// TIA Portal V19 export
// export: Created 2026-10-15T10:10:35.0564557Z, ExportSetting WithDefaults, DisplayName Totally Integrated Automation Portal, DisplayVersion V19, DisplayName TIA Portal Openness, DisplayVersion V19, DisplayName TIA Portal Version Control Interface, DisplayVersion V19, DisplayName STEP 7 Professional, DisplayVersion V19, DisplayName STEP 7 Safety, DisplayVersion V19, DisplayName WinCC Basic/Comfort/Advanced, DisplayVersion V19, DisplayName WinCC Unified, DisplayVersion V19
FUNCTION "ROLL_ShowRecipe" : Void   // FC11, SCL
{ S7_Optimized_Access := 'TRUE' }
VERSION : 0.1
// stored: AutoNumber true, IsIECCheckEnabled false, SetENOAutomatically false, UDAEnableTagReadback false
BEGIN

   "ROLL_HMI".CurrentProgram := "ROLL_State".CurrentProgram;
   "ROLL_HMI".SelectedProgram := "ROLL_State".CurrentProgram;
   "ROLL_HMI".Dwell1Seconds := "ROLL_DecodeBCD"(Value := "ROLL_DB205".DW[5]);
   "ROLL_HMI".Drain1Seconds := "ROLL_DecodeBCD"(Value := "ROLL_DB205".DW[9]);
   "ROLL_HMI".Dwell2Seconds := "ROLL_DecodeBCD"(Value := "ROLL_DB205".DW[17]);
   "ROLL_HMI".Drain2Seconds := "ROLL_DecodeBCD"(Value := "ROLL_DB205".DW[21]);
   "ROLL_HMI".Dwell3Seconds := "ROLL_DecodeBCD"(Value := "ROLL_DB205".DW[25]);
   "ROLL_HMI".Drain3Seconds := "ROLL_DecodeBCD"(Value := "ROLL_DB205".DW[29]);
   "ROLL_HMI".Dry4Seconds := "ROLL_DecodeBCD"(Value := "ROLL_DB205".DW[33]);
   "ROLL_HMI".Ultrasound1 := "ROLL_DB205".DW[13] = W#16#0001;
   "ROLL_HMI".BasketMotion := WORD_TO_INT("ROLL_DB205".DW[37]);
   "ROLL_HMI".BathLift := "ROLL_DB205".DW[41] = W#16#0001;
END_FUNCTION
